% RSLogix 500 project CTU_CTD_together.RSS, saved by version 8.30.00.16 %
PROJECT "UNTITLED"    % processor: MicroLogix 1000 %

PROGRAM FILES
  LAD 2 "MAIN_PROG"  9 rungs
  LAD 3 "USER_FAULT"  1 rungs
  LAD 4 "HSC_INT"  1 rungs
  LAD 5 "STI_INT"  1 rungs
  LAD 6, 7, 8, 9, 10, 11, 12, 13, 14, 15, 16: only END

DATA FILES
  O0 OUTPUT  5 elements
  I1 INPUT  8 elements
  S2 STATUS  33 elements
  B3 BINARY  32 elements
  T4 TIMER  40 elements
  C5 COUNTER  32 elements
  R6 CONTROL  16 elements
  N7 INTEGER  105 elements

LADDER 2 "MAIN_PROG"
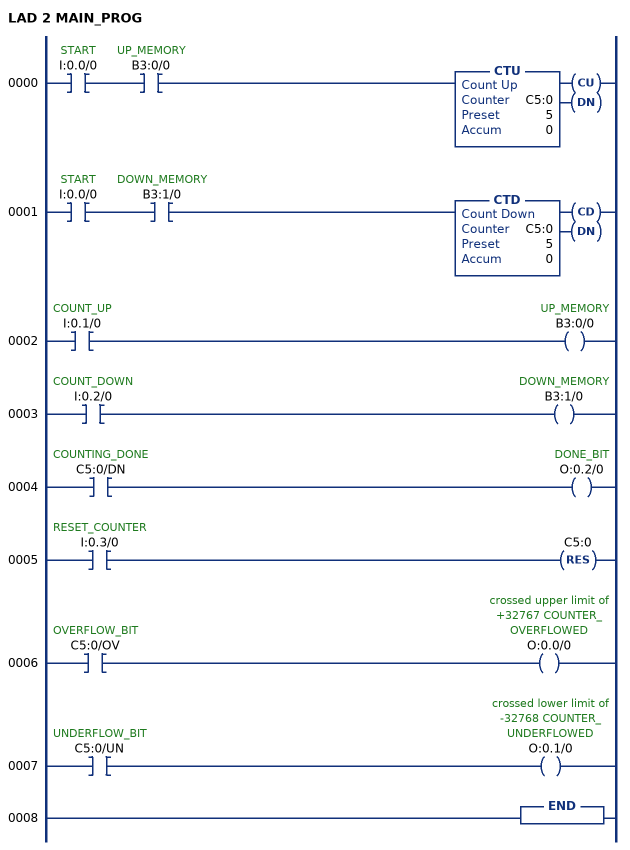
% Rung: 0 %
SOR XIC I:0.0/0 XIC B3:0/0 CTU C5:0 5 0 EOR
%   I:0.0/0  START %
%   B3:0/0  UP_MEMORY %
% Rung: 1 %
SOR XIC I:0.0/0 XIC B3:1/0 CTD C5:0 5 0 EOR
%   I:0.0/0  START %
%   B3:1/0  DOWN_MEMORY %
% Rung: 2 %
SOR XIC I:0.1/0 OTE B3:0/0 EOR
%   I:0.1/0  COUNT_UP %
%   B3:0/0  UP_MEMORY %
% Rung: 3 %
SOR XIC I:0.2/0 OTE B3:1/0 EOR
%   I:0.2/0  COUNT_DOWN %
%   B3:1/0  DOWN_MEMORY %
% Rung: 4 %
SOR XIC C5:0/DN OTE O:0.2/0 EOR
%   C5:0/DN  COUNTING_DONE %
%   O:0.2/0  DONE_BIT %
% Rung: 5 %
SOR XIC I:0.3/0 RES C5:0 EOR
%   I:0.3/0  RESET_COUNTER %
% Rung: 6 %
SOR XIC C5:0/OV OTE O:0.0/0 EOR
%   C5:0/OV  OVERFLOW_BIT %
%   O:0.0/0  COUNTER_OVERFLOWED  "crossed upper limit of +32767" %
% Rung: 7 %
SOR XIC C5:0/UN OTE O:0.1/0 EOR
%   C5:0/UN  UNDERFLOW_BIT %
%   O:0.1/0  COUNTER_UNDERFLOWED  "crossed lower limit of -32768" %
% Rung: 8 %
SOR END EOR

OTHER DOCUMENTED ADDRESSES
  I:0.0/1  COUNTINUE_COUNTING

DATA TABLE (non-zero values as saved)
DATA C5
% .PRE .ACC %
% C5:0 % 5 0
